{attribute 'qualified_only'}
{attribute 'strict'}
{attribute 'to_string'}
TYPE E_ActuatorTarget :
(
    None      := 0,     // no move commanded yet; what the outputs do is up to the actuator
    Extended  := 10,
    Retracted := 20
);
END_TYPE

(* stored: Version 1.1.0.1
   DUT E_ActuatorTarget: Id {93a96b1e-b0af-4641-b56a-2a2bb3c3ddbb} *)
